(* PLC project MixTank_MT01, Siemens AG TIA Portal V18 Update 2 *)
(* stored: creationDateTime 2025-02-11T07:52:30, contentDescription MixTank_MT01, modificationDateTime 2025-02-11T07:52:30 *)

FUNCTION FC_ScaleAnalog : REAL
  VAR_INPUT
    Raw : INT;  (* Raw analog word *)
    LoEng : REAL;
    HiEng : REAL;
  END_VAR
  VAR_TEMP
    Norm : REAL;
  END_VAR

            // 4-20 mA input on SM 1231 AI, scaled to engineering units
IF #Raw < 0 THEN
    #FC_ScaleAnalog := #LoEng;
    RETURN;
END_IF;
#Norm := NORM_X(MIN := 0, VALUE := #Raw, MAX := 32767);
#FC_ScaleAnalog := SCALE_X(MIN := #LoEng, VALUE := #Norm, MAX := #HiEng);
          
END_FUNCTION

FUNCTION_BLOCK FB_Mixer
  VAR
    Level_Pct : REAL;  (* Tank level, % *)
    Temp_C : REAL;  (* Product temperature, °C *)
    S_Heat : BOOL;  (* Step: heat *)
  END_VAR

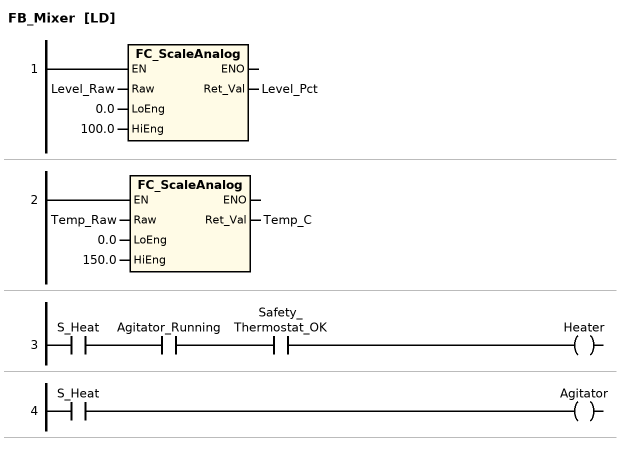
(* LD diagram, written out as Structured Text *)
Level_Pct := FC_ScaleAnalog(Level_Raw, 0.0, 100.0);
Temp_C := FC_ScaleAnalog(Temp_Raw, 0.0, 150.0);
Heater := S_Heat AND Agitator_Running AND Safety_Thermostat_OK;
Agitator := S_Heat;
END_FUNCTION_BLOCK

CONFIGURATION PLC_1
  RESOURCE CPU_1214C ON PLC
    VAR_GLOBAL  (* PLC_Tags *)
      Start_PB AT %IX0.0 : BOOL;  (* Start pushbutton (NO) *)
      Stop_PB AT %IX0.1 : BOOL;  (* Stop pushbutton (NC, TRUE = not pressed) *)
      Agitator_Running AT %IX0.4 : BOOL;  (* Agitator contactor feedback *)
      Safety_Thermostat_OK AT %IX0.5 : BOOL;  (* Safety thermostat healthy *)
      Level_Raw AT %IW96 : INT;  (* Tank level 4-20 mA *)
      Temp_Raw AT %IW98 : INT;  (* Product temperature 4-20 mA *)
      Agitator AT %QX0.0 : BOOL;  (* Agitator motor contactor *)
      Heater AT %QX0.1 : BOOL;  (* Heater contactor *)
    END_VAR
    TASK Main(INTERVAL := T#10ms, PRIORITY := 1);
    PROGRAM Mixer_DB WITH Main : FB_Mixer;
  END_RESOURCE
END_CONFIGURATION
